// Statut de l'action d'un objet (docs/04 § 5)
{attribute 'qualified_only'}
{attribute 'strict'}
TYPE E_ActStatus :
(
    Idle := 0,
    Busy := 1,
    Done := 2,
    Error := 3
) USINT;
END_TYPE

(* stored: Version 1.1.0.1, ProductVersion 3.1.4024.12
   DUT E_ActStatus: Id {71437d3f-21a8-585c-b87c-47cc968a9f15} *)
